# EPICS autosave request: 1.5.0/debian-12/7.0.10/modules/ADCore-ee039d2/db/NDCodec_settings.req
$(P)$(R)Mode
$(P)$(R)Compressor
$(P)$(R)JPEGQuality
$(P)$(R)ZlibCLevel
$(P)$(R)BloscCompressor
$(P)$(R)BloscCLevel
$(P)$(R)BloscShuffle
$(P)$(R)BloscNumThreads
$(P)$(R)LZ4HDF5BlockSize
file "NDPluginBase_settings.req", P=$(P), R=$(R)
